// TIA Portal V20 export
// export: Created 2026-10-19T18:05:22.2221153Z, ExportSetting WithDefaults, DisplayName Totally Integrated Automation Portal, DisplayVersion V20 Update 6, DisplayName TIA Portal Openness, DisplayVersion V20 Update 6, DisplayName TIA Portal Version Control Interface, DisplayVersion V20 Update 6, DisplayName SINAMICS Startdrive Advanced, DisplayVersion V20 SP1, DisplayName SINAMICS Startdrive G130, G150, S120, S150, SINAMICS MV, G220, S200, S210, DisplayVersion V20 SP1, DisplayName SINAMICS Startdrive G110M, G120, G120C, G120D, G120P, G115D, DisplayVersion V20 SP1, DisplayName STEP 7 Professional, DisplayVersion V20 Update 6, DisplayName STEP 7 Safety, DisplayVersion V20 Update 2, DisplayName WinCC Basic/Comfort/Advanced, DisplayVersion V20 Update 6, DisplayName WinCC Unified, DisplayVersion V20 Update 6
FUNCTION_BLOCK "Shuttle_TCP_Comms_Shuttle3"   // FB24, SCL
{ S7_Optimized_Access := 'TRUE' }
VERSION : 0.1
// stored: AutoNumber true, IsIECCheckEnabled false, IsRetainMemResEnabled false, MemoryReserve 100, SetENOAutomatically false, UDAEnableTagReadback false
   VAR_INPUT
      Enable : Bool;
      TCP_Configuration : "LCom_typeConfig";
   END_VAR
   VAR_OUTPUT
      Connected : Bool;
      Busy : Bool;
      Status : Word;
      Error : Bool;
   END_VAR
   VAR_IN_OUT
      TCP_Diag : "LCom_typeDiagnostics";
   END_VAR
   VAR
      SendBuffer { ExternalAccessible := 'False'; ExternalVisible := 'False'; ExternalWritable := 'False'} : Array[0..1] of Byte;
      ReceiveBuffer { ExternalAccessible := 'False'; ExternalVisible := 'False'; ExternalWritable := 'False'} : Array[0..1] of Byte;
      Send : Bool;
      SendDataLength : USInt := 2;
      Sending : Bool;
   END_VAR
BEGIN
   IF "Global_Estop" THEN
       #SendBuffer[0] := 83;
       IF NOT #Send THEN
           #Send := TRUE;
       END_IF;
   ELSE
       #SendBuffer[0] := 0;
   END_IF;

   "LCom_Communication_Shuttle3_DB"(enable := #Enable,
                                    send := #Send,
                                    sendDataLength := #SendDataLength,
                                    readDataLength := 16#FFFF_FFFF,
                                    configuration := #TCP_Configuration,
                                    connected => #Connected,
                                    sending => #Sending,
                                    busy => #Busy,
                                    error => #Error,
                                    status => #Status,
                                    sendBuffer := #SendBuffer,
                                    receiveBuffer := #ReceiveBuffer,
                                    diagnostics := #TCP_Diag);

   #SendBuffer[1] := UINT_TO_BYTE("Control_DB".VTD_Control.Current_Level);

   "Control_DB".Shuttles_Position[3].Charging := "Shuttle_MQTT_DB".Shuttle_MQTT[3].Message.Shuttle_Status.Paused;

   IF #Send AND NOT #Sending THEN
       #Send := FALSE;
   END_IF;

   IF NOT #Send THEN
       "TCP_Send_Timer_DB".TON(IN := TRUE,
                               PT := T#500ms);
   END_IF;

   IF "TCP_Send_Timer_DB".Q THEN
       #Send := TRUE;
       "TCP_Send_Timer_DB".TON(IN := FALSE,
                               PT := T#0ms);
   END_IF;
END_FUNCTION_BLOCK
